(* PLC project probe.project, CODESYS CODESYS V3.5 SP17 Patch 3 *)
(* stored: creationDateTime 2026-10-20T03:54:26.8379796, modificationDateTime 1601-01-01T03:00:00 *)

PROGRAM PRG_ProbeSfc
  VAR_INPUT
    xA : BOOL;
    xB : BOOL;
    xNext : BOOL;
  END_VAR
  VAR_OUTPUT
    iN : INT;
    xS : BOOL;
    iP : INT;
    iInit : INT;
  END_VAR

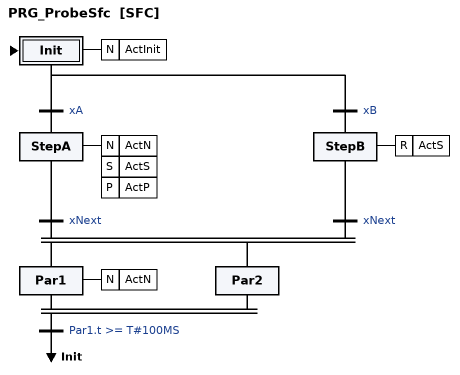
INITIAL_STEP Init:
  ActInit(N);
END_STEP
TRANSITION FROM Init TO StepA
  := xA;
END_TRANSITION
TRANSITION FROM Init TO StepB
  := xB;
END_TRANSITION
STEP StepA:
  ActN(N);
  ActS(S);
  ActP(P);
END_STEP
TRANSITION FROM StepA TO (Par1, Par2)
  := xNext;
END_TRANSITION
STEP StepB:
  ActS(R);
END_STEP
TRANSITION FROM StepB TO (Par1, Par2)
  := xNext;
END_TRANSITION
STEP Par1:
  ActN(N);
END_STEP
TRANSITION FROM (Par1, Par2) TO Init
  := Par1.t >= T#100MS;
END_TRANSITION
STEP Par2:
END_STEP

ACTION ActInit:
                iInit := iInit + 1;

              
END_ACTION

ACTION ActN:
                iN := iN + 1;

              
END_ACTION

ACTION ActS:
                xS := TRUE;

              
END_ACTION

ACTION ActP:
                iP := iP + 1;

              
END_ACTION
END_PROGRAM
